// TIA Portal V21 export
ORGANIZATION_BLOCK "Parallel"   // OB1, LAD
BEGIN

REGION Network 1: Seal-in
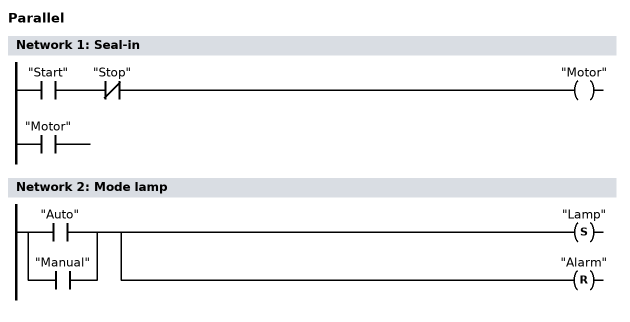
   "Motor" := "Start" AND NOT "Stop";
END_REGION

REGION Network 2: Mode lamp
   RUNG wire#powerrail
      Contact( "Auto" )
      wire#w1
      S_Coil( "Lamp" )
   END_RUNG
   RUNG wire#powerrail
      Contact( "Manual" )
   END_RUNG wire#w1
   RUNG wire#w1
      R_Coil( "Alarm" )
   END_RUNG
   // the same network as SCL:
   IF "Auto" OR "Manual" THEN
       "Lamp" := TRUE;
       "Alarm" := FALSE;
   END_IF;
END_REGION
END_ORGANIZATION_BLOCK
